FUNCTION_BLOCK FillRetry_AOI (* Migrated from IEC 61131-3 ST *)
  (* Standard: 61499-2 *)
  (* Version 1.0, 2026-11-06, st2fb *)
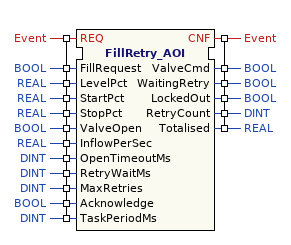
  EVENT_INPUT
    REQ WITH FillRequest, LevelPct, StartPct, StopPct, ValveOpen, InflowPerSec, OpenTimeoutMs, RetryWaitMs, MaxRetries, Acknowledge, TaskPeriodMs;
  END_EVENT
  EVENT_OUTPUT
    CNF WITH ValveCmd, WaitingRetry, LockedOut, RetryCount, Totalised;
  END_EVENT
  VAR_INPUT
    FillRequest : BOOL;
    LevelPct : REAL;
    StartPct : REAL;
    StopPct : REAL;
    ValveOpen : BOOL;
    InflowPerSec : REAL;
    OpenTimeoutMs : DINT;
    RetryWaitMs : DINT;
    MaxRetries : DINT;
    Acknowledge : BOOL;
    TaskPeriodMs : DINT;
  END_VAR
  VAR_OUTPUT
    ValveCmd : BOOL;
    WaitingRetry : BOOL;
    LockedOut : BOOL;
    RetryCount : DINT;
    Totalised : REAL;
  END_VAR
  VAR
    Demand : BOOL := FALSE;
    WaitActive : BOOL := FALSE;
    OpenTimer_TimerEnable : BOOL := FALSE;
    OpenTimer_PRE : DINT := 0;
    OpenTimer_EN : BOOL := FALSE;
    OpenTimer_TT : BOOL := FALSE;
    OpenTimer_DN : BOOL := FALSE;
    OpenTimer_ACC : DINT := 0;
    WaitTimer_TimerEnable : BOOL := FALSE;
    WaitTimer_PRE : DINT := 0;
    WaitTimer_EN : BOOL := FALSE;
    WaitTimer_TT : BOOL := FALSE;
    WaitTimer_DN : BOOL := FALSE;
    WaitTimer_ACC : DINT := 0;
    Retries_CUEnable : BOOL := FALSE;
    Retries_PRE : DINT := 0;
    Retries_ACC : DINT := 0;
    Retries_DN : BOOL := FALSE;
    Retries_PREV : BOOL := FALSE;
    AckOneShot_InputBit : BOOL := FALSE;
    AckOneShot_OutputBit : BOOL := FALSE;
    AckOneShot_PREV : BOOL := FALSE;
    OpenTimer_PREV : BOOL := FALSE;
    WaitTimer_PREV : BOOL := FALSE;
  END_VAR
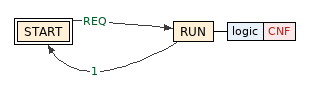
  EC_STATES
    START;
    RUN : logic -> CNF;
  END_STATES
  EC_TRANSITIONS
    START TO RUN := REQ;
    RUN TO START := 1;
  END_TRANSITIONS
  ALGORITHM logic IN ST:
IF LevelPct <= StartPct THEN
  Demand := TRUE;
ELSIF LevelPct >= StopPct THEN
  Demand := FALSE;
END_IF;

Retries_CUEnable := OpenTimer_DN;
Retries_PRE := MaxRetries;
IF Retries_CUEnable AND NOT Retries_PREV THEN
  Retries_ACC := Retries_ACC + 1;
END_IF;
Retries_PREV := Retries_CUEnable;
Retries_DN := Retries_ACC >= Retries_PRE;
RetryCount := Retries_ACC;
LockedOut := Retries_DN;

IF OpenTimer_DN AND NOT LockedOut THEN
  WaitActive := TRUE;
END_IF;
WaitTimer_TimerEnable := WaitActive;
WaitTimer_PRE := RetryWaitMs;
WaitTimer_EN := WaitTimer_TimerEnable;
IF WaitTimer_EN THEN
  IF WaitTimer_PREV AND NOT WaitTimer_DN THEN
    WaitTimer_ACC := WaitTimer_ACC + TaskPeriodMs;
    IF WaitTimer_ACC >= WaitTimer_PRE THEN
      WaitTimer_ACC := WaitTimer_PRE;
      WaitTimer_DN := TRUE;
    END_IF;
  END_IF;
ELSE
  WaitTimer_ACC := 0;
  WaitTimer_DN := FALSE;
END_IF;
WaitTimer_TT := WaitTimer_EN AND NOT WaitTimer_DN;
WaitTimer_PREV := WaitTimer_EN;
WaitingRetry := WaitTimer_TT;
IF WaitTimer_DN THEN
  WaitActive := FALSE;
END_IF;

ValveCmd := FillRequest AND Demand AND NOT LockedOut AND NOT WaitActive;

OpenTimer_TimerEnable := ValveCmd AND NOT ValveOpen;
OpenTimer_PRE := OpenTimeoutMs;
OpenTimer_EN := OpenTimer_TimerEnable;
IF OpenTimer_EN THEN
  IF OpenTimer_PREV AND NOT OpenTimer_DN THEN
    OpenTimer_ACC := OpenTimer_ACC + TaskPeriodMs;
    IF OpenTimer_ACC >= OpenTimer_PRE THEN
      OpenTimer_ACC := OpenTimer_PRE;
      OpenTimer_DN := TRUE;
    END_IF;
  END_IF;
ELSE
  OpenTimer_ACC := 0;
  OpenTimer_DN := FALSE;
END_IF;
OpenTimer_TT := OpenTimer_EN AND NOT OpenTimer_DN;
OpenTimer_PREV := OpenTimer_EN;

IF ValveCmd AND ValveOpen THEN
  Totalised := Totalised + InflowPerSec * DINT_TO_REAL(TaskPeriodMs) / 1000.0;
END_IF;

AckOneShot_InputBit := Acknowledge;
AckOneShot_OutputBit := AckOneShot_InputBit AND NOT AckOneShot_PREV;
AckOneShot_PREV := AckOneShot_InputBit;
IF AckOneShot_OutputBit THEN
  Retries_ACC := 0;
  Retries_DN := FALSE;
  OpenTimer_ACC := 0;
  OpenTimer_EN := FALSE;
  OpenTimer_TT := FALSE;
  OpenTimer_DN := FALSE;
  OpenTimer_PREV := FALSE;
  WaitTimer_ACC := 0;
  WaitTimer_EN := FALSE;
  WaitTimer_TT := FALSE;
  WaitTimer_DN := FALSE;
  WaitTimer_PREV := FALSE;
  WaitActive := FALSE;
END_IF;
  END_ALGORITHM
END_FUNCTION_BLOCK
